Fanuc KAREL source: kt00870.KL

PROGRAM KT00870
%NOLOCKGROUP
VAR
R1:REAL;R2:REAL;OUT:INTEGER
BEGIN
--
--
R1=2.0
R2=3.0
R1=2.0
R2=3.0
OUT=TRUNC(R1)
END KT00870
